Universal Robots PolyScope program: P1140 INVITE_training_1.urp

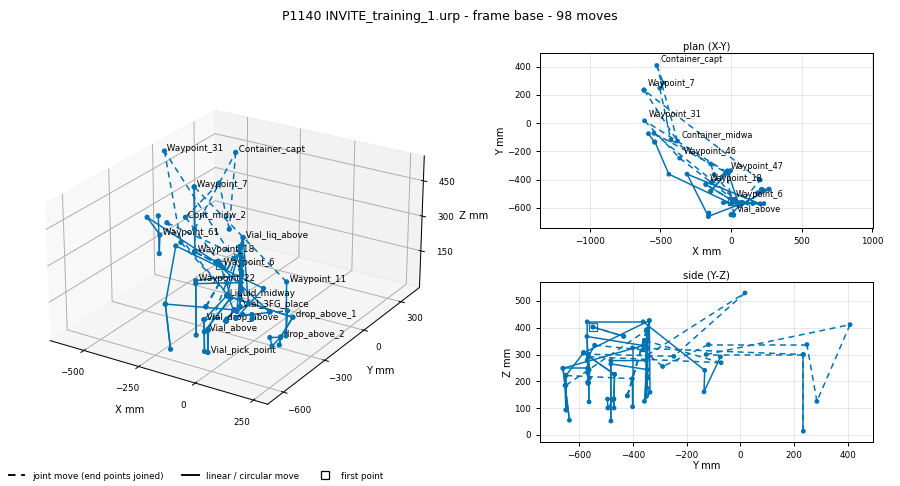
[picture p0: tool path of P1140 INVITE_training_1.urp in frame base, 98 of 125 moves have a stored position in this frame; points joined in program order, loops and branches not executed]
Program P1140 INVITE_training_1 (installation=default directory=/programs/02 Main Routines createdIn=5.10.1 lastSavedIn=5.19.0 robotSerialNumber=20245590068)
Calibrated DH parameters: a=[0.00013, -0.03651, -0.389144, 0.000102, 0.000008, 0]; d=[0.162613, 192.230671, -179.915756, -12.181517, 0.099698, 0.099535]; alpha=[1.57038, 0.002205, 0.004138, 1.570804, -1.571025, 0]; deltaTheta=[-0.000001, 1.484886, 4.928506, -0.130209, 0, 0]
InitVariablesNode variables(variable(name=AMR_Position, expression=struct(position_identifier=0, x1=0, x2=0, y1=0, y2=0, theta1=0, theta2=0)), variable(name=CAM_Pose, expression=p[0,0,0,0,0,0]), variable(name=CAM_Relation, expression=""), variable(name=CMD_Abort, expression=False), variable(name=CMD_Clear, expression=False), variable(name=CMD_Reset, expression=False), variable(name=CMD_Start, expression=False), variable(name=CMD_Suspend, expression=False), variable(name=CMD_Unhold, expression=False), variable(name=CMD_Unsuspend, expression=False), variable(name=CNT_Rack_Output, expression=0), variable(name=FNC_Freedrive, expression=False), variable(name=PRC_TubCounter, expression=0), variable(name=PRC_TubNumber, expression=0), variable(name=STP, expression=0), variable(name=TMR_Barcode, expression=0), variable(name=easyPickCount, expression=0), variable(name=easyPickCount_1, expression=0), variable(name=easyPickCount_2, expression=0), variable(name=easyPickCount_3, expression=0), variable(name=easyPickNoObj, expression=0), variable(name=easyPickNoObj_1, expression=0), variable(name=easyPickNoObj_2, expression=0), variable(name=easyPickNoObj_3, expression=0), variable(name=easyPickParts, expression=0), variable(name=easyPickParts_1, expression=0), variable(name=easyPickParts_2, expression=0), variable(name=easyPickParts_3, expression=0))
BeforeStart
  Folder Scripts
    Script file /programs/04 Scripts/001 SCRIPT Errors and Warnings Deifnes V0.2.script
      | #*****************************************************
      | # customer          :   UK Essen
      | # project name      :   P1132
      | #****************************************************
      | # controller        :
      | # software          :
      | #****************************************************
      | # author            :   E.Petrichenko
      | # Copyright (c)     :   United Robotics Group Health and Food GmbH
      | #                       An der Riede 2
      | #                       28816 Stuhr
      | #                       Germany
      | #****************************************************
      | # description       :   centrifuge actions for the application
      | # version:      	:   0.1
      | # created           :   22.08.2024
      | # updated           :
      | #****************************************************
      | # modifications     :
      | #
      | # date              :
      | # name              :
      | # reason            :
      | #****************************************************
      | 
      | 
      | #################################### VARIABLES DEFINITIONS ###################################
      | 
      | ERROR_POSE_NOT_REACHABLE = 1002
      | ERROR_ROBOT_ARM_NOT_IN_HOME_POSE = 1006
      | ERROR_NO_OBJECT_TO_PICK = 1010
      | ERROR_NOT_DOCKED = 2003
      | ERROR_NOT_REACHABLE_TARGET = 2007
      | ERROR_CHARGING_NOT_STARTED = 2008
      | ERROR_AMR_WRONG_MODE = 2009
      | ERROR_UNKNOWN_POSE = 2010
      | ERROR_NO_LANDMARK = 3002
      | ERROR_WRONG_ORDER = 4002
      | ERROR_CENTRIFUGE_CONNECTION = 5001
      | ERROR_CENTRIFUGE_POWER = 5002
      | ERROR_CENTRIFUGE = 5003
      | ERROR_CENTRIFUGE_LID = 5004
      | ERROR_CANNOT_OPEN_HATCH = 5006
      | ERROR_CANNOT_CLOSE_HATCH = 5008
      | ERROR_CANNOT_ROTATE = 5010
      | ERROR_CANNOT_START = 5011
      | ERROR_WRONG_KEY_POSE = 5012
      | ERROR_MISSIING_CENTRACK = 5013
      | 
      | WARNING_POSE_NOT_REACHABLE = 1002
      | WARNING_BATTERY_LEVEL = 2002
      | WARNING_NOT_REACHABLE_TARGET = 2007
      | 
      | 
      | ERROR = struct(
      |     FLAG = False,
      |     ID = 0,
      |     MSG = "")
      | 
      | WARNING = struct(
      |     FLAG = False,
      |     ID = 0,
      |     MSG = "")
      | 
      | 
      | #################################### FUNCTIONS ###################################
      | 
      | def set_error(error_id):
      |     ERROR.ID = error_id
      |     if (ERROR.ID == 0):
      |         ERROR.FLAG = False
      |         ERROR.MSG = ""
      |     else:
      |         ERROR.FLAG = True
      |         if(ERROR.ID == ERROR_POSE_NOT_REACHABLE):
      |             ERROR.MSG = "Pose is not reachable"
      |         elif(ERROR.ID == ERROR_NO_OBJECT_TO_PICK):
      |             ERROR.MSG = "No object to pick"
      |         elif(ERROR.ID == ERROR_NO_LANDMARK):
      |             ERROR.MSG = "No landmark detected"
      |         elif(ERROR.ID == ERROR_ROBOT_ARM_NOT_IN_HOME_POSE):
      |             ERROR.MSG = "Robot arm cannot go to home pose"
      |         elif(ERROR.ID == ERROR_AMR_WRONG_MODE):
      |             ERROR.MSG = "AMR is in the wrong mode"
      |         elif(ERROR.ID == ERROR_NOT_DOCKED):
      |             ERROR.MSG = "Could not dock to the charger"
      |         elif(ERROR.ID == ERROR_NOT_REACHABLE_TARGET):
      |             ERROR.MSG = "Could not reach the target"
      |         elif(ERROR.ID == ERROR_CHARGING_NOT_STARTED):
      |             ERROR.MSG = "Could not start charging"
      |         elif(ERROR.ID == ERROR_UNKNOWN_POSE):
      |             ERROR.MSG = "Unknown navigation target"
      |         elif(ERROR.ID == ERROR_CANNOT_OPEN_HATCH):
      |             ERROR.MSG = "Centrifuge Cannot open the hatch"
      |         elif(ERROR.ID == ERROR_CENTRIFUGE_CONNECTION):
      |             ERROR.MSG = "Cannot reach centrifuge"
      |         elif (ERROR.ID == ERROR_CANNOT_CLOSE_HATCH):
      |             ERROR.MSG = "Centrifuge Cannot close the hatch"
      |         elif (ERROR.ID == ERROR_CANNOT_START):
      |             ERROR.MSG = "Centrifuge Cannot start"
      |         elif (ERROR.ID == ERROR_CANNOT_ROTATE):
      |             ERROR.MSG = "Centrifuge Cannot rotate the rotor"
      |         elif (ERROR.ID == ERROR_WRONG_ORDER):
      |             ERROR.MSG = "Wrong parameter was recieved"
      |         elif (ERROR.ID == ERROR_CENTRIFUGE):
      |             ERROR.MSG = "Centrifuge is in Error"
      |         elif (ERROR.ID == ERROR_WRONG_KEY_POSE):
      |             ERROR.MSG = "Key is in the wrong position"
      |         elif(ERROR.ID == ERROR_MISSIING_CENTRACK):
      |             ERROR.MSG = "Missing rack for centrifuge set"
      |         elif(ERROR.ID == ERROR_CENTRIFUGE_POWER):
      |             ERROR.MSG = "Centrifuge is turned off"
      |         elif(ERROR.ID == ERROR_CENTRIFUGE_LID):
      |             ERROR.MSG = "Lid of the centrifuge is opened"
      |         else:
      |             ERROR.MSG = "Unknown code"
      |         end
      |         textmsg("ERROR:",ERROR)
      |     end
      | end
      | 
      | def set_warning(warning_id):
      |     WARNING.ID = warning_id
      |     if (WARNING.ID == 0):
      |         WARNING.FLAG = False
      |         WARNING.MSG = ""
      |     else:
      |         WARNING.FLAG = True
      |         if(WARNING.ID == WARNING_POSE_NOT_REACHABLE):
      |             WARNING.MSG = "Pose is not reachable"
      |         elif(WARNING.ID == WARNING_BATTERY_LEVEL):
      |             WARNING.MSG = "Batery level dropped to a certain level"
      |         elif(WARNING.ID == WARNING_NOT_REACHABLE_TARGET):
      |             WARNING.MSG = "Not reachable location of AMR"
      |         else:
      |             WARNING.MSG = "Unknown code"
      |         end
      |         textmsg("WARNING:",WARNING)
      |     end
      | end
      | 
      | 
      | def reset_error():
      |   ERROR.ID = 0
      |   ERROR.FLAG = False
      |   ERROR.MSG = ""
      | end
      | 
      | 
      | def reset_warning():
      |     WARNING.ID = 0
      |     WARNING.FLAG = False
      |     WARNING.MSG = ""
      |   end
    Script file /programs/04 Scripts/SCRIPT uGO V7.11.1.script
      | #*****************************************************
      | # customer          :
      | # project name      :   Standard Application
      | #****************************************************
      | # controller        :
      | # software          :
      | #****************************************************
      | # author            :   P. Koehnke
      | # Copyright (c)     :   United Robotics Group
      | #                       An der Riede 2
      | #                       28816 Stuhr
      | #                       Germany
      | #****************************************************
      | # description       :   interface for uGo
      | # version:      	:   6.0
      | # created           :   21.04.2022
      | # updated           :
      | #****************************************************
      | # modifications     :   add new rpc-functions to interchange more data
      | #
      | # date              :   2024-02-29
      | # name              :   P. Koehnke
      | # reason            :   implemtentation of PackML behavoiur in uGO
      | #****************************************************
      | #****************************************************
      | # modifications     :   add reflecting the UID of the uGO task back to uGO
      | #
      | # date              :   2024-07-02
      | # name              :   P. Koehnke
      | # reason            :   be sure to finish the right tasks
      | #****************************************************
      | 
      | # available rpc-functions:
      | #.on('con_check', (err, _params, callback) => callback(err, this.con_check()))
      | #.on('read_input', (err, params, callback) => callback(err, this.read_input(params[0], params[1])))
      | #.on('write_output', (err, params, callback) => callback(err, this.write_output(params[0], params[1], params[2])))
      | #.on('read_status', (err, params, callback) => callback(err, this.read_status(params[0])))
      | #.on('write_status', (err, params, callback) => callback(err, this.write_status(params[0], params[1])))
      | #.on('send_template', (err, params, callback) => callback(err, this.receive_state(params[0])))
      | #.on('receive_event', (err, params, callback) => callback(err, this.send_event()))
      | #.on('send_state', (err, params, callback) => callback(err, this.receive_state(params[0])))
      | #.on('send_error', (err, params, callback) => callback(err, this.receive_error(params[0])))
      | #.on('NotFound', (methodCalled, params) => LOG.warn('Method "', methodCalled, '" does not exist. ', { params }));
      | 
      | # =======================================================================
      | local IDX_CMD_STOP = 0
      | local IDX_CMD_RESET = 1
      | local IDX_CMD_START = 2
      | local IDX_CMD_HOLD = 3
      | local IDX_CMD_UNHOLD = 4
      | local IDX_CMD_SUSPEND = 5
      | local IDX_CMD_UNSUSPEND = 6
      | local IDX_CMD_ABORT = 7
      | local IDX_CMD_CLEAR = 8
      | local IDX_FNC_FREEDRIVE = 9
      | 
      | # uGo specific declarations
      | global UGO_Request_ID = ""
      | global UGO_UNIT_Task = ""
      | global UGO_Task_ID = 0
      | global UGO_Event = ""
      | local UGO_Enable_Control = False
      | local UGO = rpc_factory("xmlrpc", "http://192.168.12.120:8080")
      | local UGO_Ctrl_Cmd = [False, False, False, False, False, False, False, False, False, False]
      | 
      | local UGO_AMR_Pos = struct(position_identifier=0, x1=0, x2=0, y1=0, y2=0, theta1=0, theta2=0)
      | local UGO_EOAT = struct(object_picked=False)
      | 
      | def ugo_init(enable=True, rpc_address="http://192.168.12.120:8080"):
      |     # connection with uGo
      |     if enable:
      |         UGO = rpc_factory("xmlrpc", rpc_address)
      |         UGO_Enable_Control = True
      |     else:
      |         UGO_Enable_Control = False
      |     end
      | end
      | 
      | def ugo_event_controller():
      |     # interpret the given command and map it to the internal commands
      |     if UGO_Enable_Control:
      |         UGO_Event = UGO.receive_event()
      |     end
      | 
      |     UGO_Ctrl_Cmd[IDX_CMD_STOP] = (UGO_Event == "stop")
      |     UGO_Ctrl_Cmd[IDX_CMD_RESET] = (UGO_Event == "reset")
      |     UGO_Ctrl_Cmd[IDX_CMD_START] = (UGO_Event == "start")
      |     UGO_Ctrl_Cmd[IDX_CMD_HOLD] = (UGO_Event == "hold")
      |     UGO_Ctrl_Cmd[IDX_CMD_UNHOLD] = (UGO_Event == "un_hold")
      |     UGO_Ctrl_Cmd[IDX_CMD_SUSPEND] = (UGO_Event == "suspend")
      |     UGO_Ctrl_Cmd[IDX_CMD_UNSUSPEND] = (UGO_Event == "un_suspend")
      |     UGO_Ctrl_Cmd[IDX_CMD_ABORT] = (UGO_Event == "abort")
      |     UGO_Ctrl_Cmd[IDX_CMD_CLEAR] = (UGO_Event == "clear")
      |     UGO_Ctrl_Cmd[IDX_FNC_FREEDRIVE] = (UGO_Event == "freedrive")
      | 
      |     return UGO_Ctrl_Cmd
      | end
      | 
      | def ugo_translate_pml_state():
      |     # translate the current PML State to a string
      |     if (STATE == 1):
      |         return "STOPPING"
      |     elif (STATE == 2):
      |         return "STOPPED"
      |     elif (STATE == 3):
      |         return "RESETTING"
      |     elif (STATE == 4):
      |         return "IDLE"
      |     elif (STATE == 5):
      |         return "STARTING"
      |     elif (STATE == 6):
      |         return "EXECUTE"
      |     elif (STATE == 7):
      |         return "COMPLETING"
      |     elif (STATE == 8):
      |         return "COMPLETE"
      |     elif (STATE == 9):
      |         return "HOLDING"
      |     elif (STATE == 10):
      |         return "HELD"
      |     elif (STATE == 11):
      |         return "UNHOLDING"
      |     elif (STATE == 12):
      |         return "SUSPENDING"
      |     elif (STATE == 13):
      |         return "SUSPENDED"
      |     elif (STATE == 14):
      |         return "UNSUSPENDING"
      |     elif (STATE == 15):
      |         return "ABORTING"
      |     elif (STATE == 16):
      |         return "ABORTED"
      |     elif (STATE == 17):
      |         return "CLEARING"
      |     else:
      |         return "UNKNOWN"
      |     end
      | end
      | 
      | def ugo_update_outputs():
      |     #Update the outputs to uGo via xmplrpc service
      |     UGO.write_status("ROB_Skill", UGO_UNIT_Task)
      |     UGO.write_status("ROB_Battery", AMR_Battery)
      |     UGO.write_status("ROB_Gripper", OBJ_Picked)
      |     UGO.send_state(ugo_translate_pml_state(), UGO_UNIT_Task)
      |     UGO.send_error(ERROR.ID)
      |     #UGO.send_position(AMR_Position)
      | end
      | 
      | def ugo_get_task():
      |     # get the actual task to work on
      |     # added: reflecting the UID of the task back to uGO
      |     UGO_UNIT_Task = UGO.read_status("DSH_Workflow")
      |     if (UGO_UNIT_Task != ""):
      |         UGO_Request_ID = str_sub(UGO_UNIT_Task, 0, 39)
      |         UGO_Task_ID = to_num(str_sub(UGO_UNIT_Task, 40, 2))
      |         #ugo_tasks()
      |         return UGO_Task_ID
      |     else:
      |         return 0
      |     end
      | end
      | 
      | def ugo_pml_stopping():
      |     return True
      | end
      | 
      | def ugo_pml_resetting():
      |     ugo_get_task()
      |     if (UGO_UNIT_Task == ""):
      |         UGO_Request_ID = ""
      |         UGO_Task_ID = 0
      |         return True
      |     end
      |     return False
      | end
      | 
      | def ugo_pml_starting():
      |     #UGO_Task_Content = UGO.receive_task()
      |     return (UGO_UNIT_Task != "")
      | end
      | 
      | def ugo_pml_holding():
      |     return True
      | end
      | 
      | def ugo_pml_unholding():
      |     return True
      | end
      | 
      | def ugo_pml_suspending():
      |     return True
      | end
      | 
      | def ugo_pml_unsuspending():
      |     return True
      | end
      | 
      | def ugo_pml_completing():
      |     return True
      | end
      | 
      | def ugo_pml_aborting():
      |     return True
      | end
      | 
      | def ugo_pml_clearing():
      |     return True
      | end
      | 
      | # =======================================================================
      | # end of uGO script
      | # =======================================================================
    SuppressedNode
      Script file /programs/04 Scripts/SCRIPT Centrifuge Actions V0.3.script
        | #*****************************************************
        | # customer          :   UK Essen
        | # project name      :   P1132
        | #****************************************************
        | # controller        :
        | # software          :
        | #****************************************************
        | # author            :   E.Petrichenko
        | # Copyright (c)     :   United Robotics Group Health and Food GmbH
        | #                       An der Riede 2
        | #                       28816 Stuhr
        | #                       Germany
        | #****************************************************
        | # description       :   centrifuge actions for the application
        | # version:      	:   0.1
        | # created           :   22.08.2024
        | # updated           :
        | #****************************************************
        | # modifications     :
        | #
        | # date              :
        | # name              :
        | # reason            :
        | #****************************************************
        | 
        | 
        | #################################### VARIABLES DEFINITIONS ###################################
        | CNT_RESET_LOAD_TIMER = 60
        | CNT_Rotate_Error = False
        | CNT_Error = ""
        | CNT_LidState = 0
        | CNT_Timer_Start = 0
        | CNT_Timer_Counting = False
        | CNT_Hatch_State = 0
        | global CNT_State_Actual  = 0
        | CNT_KeyState = 0
        | Cent=rpc_factory("xmlrpc","http://192.168.12.125:50002")
        | 
        | ACTION_OPEN_HATCH = 5
        | ACTION_CLOSE_HATCH = 6
        | ACTION_START = 9
        | ACTION_INSPECT = 16
        | ACTION_ROTATE = 23
        | 
        | CNT_STATES_INIT = struct (
        |     UNSTARTABLE = 1,
        |     STOPPED = 2,
        |     STOPPED_UNSTARTABLE = 3,
        |     RUN_UP = 4,
        |     RUNNING = 8)
        | 
        | 
        | KEY_STATE_INIT = struct (
        |     TEACH = 1,
        |     LOCKED = 2,
        |     MIDDLE = 3)
        | 
        | LID_STATE_INIT = struct (
        |     CLOSED = 0,
        |     OPENED = 1)
        | #stopped_unstartable happens when lid or hatch is open
        | 
        | #################################### THREADS ###################################
        | 
        | thread Timer_CentThread():
        |     while (True):
        |         if (CNT_Timer_Counting):
        |             CNT_Timer_Start = CNT_Timer_Start + get_steptime()
        |         end
        |         sync()
        |     end
        | end
        | thread_timer_cent = run Timer_CentThread()
        | 
        | thread Cent_Thread():
        |     while (True):
        |         CNT_Hatch_State = Cent.hatchstate()
        |         CNT_State_Actual  = Cent.state()
        |         log_hatch_state(CNT_Hatch_State)
        |         log_centrifuge_state(CNT_State_Actual)
        |         sleep(0.5)
        |     end
        | end
        | run Cent_Thread()
        | 
        | #################################### FUNCTIONS ###################################
        | 
        | 
        | 
        | def cent_error_check():
        |     CNT_Error = Cent.geterror()
        |     CNT_KeyState = Cent.keystate()
        |     CNT_LidState = Cent.lidstate()
        | 
        |     if (CNT_Error == "88888888"):
        |         set_error(ERROR_CENTRIFUGE_POWER)
        |     elif (CNT_Error != "00000000"):
        |         set_error(ERROR_CENTRIFUGE)
        |         textmsg("CNT_Error:",CNT_Error)
        |     elif (CNT_KeyState != KEY_STATE_INIT.LOCKED):
        |         set_error(ERROR_WRONG_KEY_POSE)
        |     elif (CNT_LidState == LID_STATE_INIT.OPENED):
        |       set_error(ERROR_CENTRIFUGE_LID)
        |     end
        | 
        | end
        | 
        | 
        | def execute_cent_action(cent_action, cent_slot = 0):
        | 
        |     if (cent_action == ACTION_OPEN_HATCH):
        |         local cnt_hatch_moved = 0
        |         if (CNT_State_Actual  == 2):
        |             cnt_hatch_moved = Cent.move_hatch(2)
        |             if (cnt_hatch_moved == -1):
        |                 set_error(ERROR_CANNOT_OPEN_HATCH)
        |             end
        |         elif (CNT_State_Actual  == 3):
        |             textmsg("WARNING: Centrifuge is already opened", True)
        |         else:
        |             set_error(ERROR_WRONG_ORDER)
        |             textmsg("ERROR: Centrifuge state is not corresponded with the required task", True)
        |         end
        | 
        |     elif (cent_action == ACTION_CLOSE_HATCH):
        |         cnt_hatch_moved = Cent.move_hatch(1)
        |         if (cnt_hatch_moved == -1):
        |             set_error(ERROR_CANNOT_CLOSE_HATCH)
        |         end
        | 
        |     elif (cent_action == ACTION_START):
        |         Cent.start()
        |         CNT_Timer_Start = 0
        |         CNT_Timer_Counting = True
        |         while ((CNT_State_Actual  != CNT_STATES_INIT.RUN_UP and CNT_State_Actual  != CNT_STATES_INIT.RUNNING) and CNT_Timer_Start < CNT_RESET_LOAD_TIMER and not CMD_Stop and not CMD_Hold):
        |             sleep(0.5)
        | 
        |         end
        | CNT_Timer_Counting = False
        |         if (CNT_Timer_Start >= CNT_RESET_LOAD_TIMER ):
        |             set_error(ERROR_CANNOT_START)
        |             if (CNT_State_Actual == CNT_STATES_INIT.UNSTARTABLE or CNT_State_Actual == CNT_STATES_INIT.STOPPED_UNSTARTABLE):
        |                 set_error(ERROR_WRONG_ORDER)
        |                 textmsg("ERROR: Centrifuge state is not corresponded with the required task", True)
        |             end
        |         end
        |     elif (cent_action == ACTION_INSPECT):
        |         if (CNT_Rotate_Error == False):
        |             set_error(ERROR_CANNOT_ROTATE)
        |         else:
        |             CNT_Rotate_Error = Cent.posreached(6 *(cent_slot-1) + 1)
        |             if (CNT_Rotate_Error == False):
        |               set_error(ERROR_CANNOT_ROTATE)
        |             end
        |         end
        | 
        | 
        |     elif (cent_action == ACTION_ROTATE):
        |         CNT_Rotate_Error = False
        |         CNT_Rotate_Error = Cent.move_rotor(6 *(cent_slot-1) + 1)
        |         return CNT_Rotate_Error
        |     else:
        |         set_error(ERROR_WRONG_ORDER)
        |     end
        | end
    Script file /programs/04 Scripts/SCRIPT PackML V1.2.1.script
      | # PackML
      | 
      | IO_ADDRESS_CMD_STOP = 1
      | IO_ADDRESS_CMD_RESET = 7
      | IO_ADDRESS_CMD_START = 0
      | 
      | EXT_ADDRESS_CMD_STOP = 0
      | EXT_ADDRESS_CMD_RESET = 1
      | EXT_ADDRESS_CMD_START = 2
      | EXT_ADDRESS_CMD_HOLD = 3
      | EXT_ADDRESS_CMD_UNHOLD = 4
      | EXT_ADDRESS_CMD_SUSPEND = 5
      | EXT_ADDRESS_CMD_UNSUSPEND = 6
      | EXT_ADDRESS_CMD_ABORT = 7
      | EXT_ADDRESS_CMD_CLEAR = 8
      | EXT_ADDRESS_FNC_FREEDRIVE = 9
      | 
      | global EXT_CtrlCmd = [False, False, False, False, False, False, False, False, False, False]
      | 
      | EXT_Control_by = "uGO"
      | 
      | global CMD_Abort = False
      | global CMD_Clear = False
      | global CMD_Stop = False
      | global CMD_Reset = False
      | global CMD_Start = False
      | global CMD_Hold = False
      | global CMD_Unhold = False
      | global CMD_Suspend = False
      | global CMD_Unsuspend = False
      | global FNC_Freedrive = False
      | 
      | CND_Suspend = False         # condition for suspend command
      | CND_Unsuspend = False       # condition for unsuspend command
      | 
      | thread Get_Pml_Command():
      |     while (True):
      |         if (EXT_Control_by == "uGO"):
      |             EXT_CtrlCmd = ugo_event_controller()
      |         elif (EXT_Control_by == "Leitsystem"):
      |             # EXT_CtrlCmd = Leitsystem
      |         end
      |         # ---------- Abort ---------- #
      |         if ((not STATE == 15) and (not STATE == 16) and EXT_CtrlCmd[EXT_ADDRESS_CMD_ABORT]):
      |             CMD_Abort = True
      |             CMD_Stop = False
      |         elif ((STATE == 17) and not EXT_CtrlCmd[EXT_ADDRESS_CMD_ABORT]):
      |             CMD_Abort = False
      |         end
      |         # ---------- Stop ---------- #
      |         if ((not STATE == 1) and (not STATE == 2) and (get_standard_digital_in(IO_ADDRESS_CMD_STOP) or EXT_CtrlCmd[EXT_ADDRESS_CMD_STOP])):
      |             CMD_Stop = True
      |             if get_standard_digital_in(IO_ADDRESS_CMD_STOP):
      |                 log_state("Stop command by pushbutton")
      |             elif EXT_CtrlCmd[EXT_ADDRESS_CMD_STOP]:
      |                 log_state("Stop command by external control")
      |             end
      |         elif (STATE == 2) and (not get_standard_digital_in(IO_ADDRESS_CMD_STOP)) and (not EXT_CtrlCmd[EXT_ADDRESS_CMD_STOP]):
      |             CMD_Stop = False
      |         end
      |         CMD_Hold = (STATE == 6 or STATE == 10) and not CMD_Stop and (ERROR.FLAG or EXT_CtrlCmd[EXT_ADDRESS_CMD_HOLD])
      |         CMD_Reset = (STATE == 2 or STATE == 8) and not CMD_Stop and (read_input_boolean_register(5) or EXT_CtrlCmd[EXT_ADDRESS_CMD_RESET])
      |         CMD_Start = (STATE == 4) and not CMD_Stop and (get_standard_digital_in(IO_ADDRESS_CMD_START) or EXT_CtrlCmd[EXT_ADDRESS_CMD_START])
      |         CMD_Unhold = (STATE == 10) and not CMD_Stop and (get_standard_digital_in(IO_ADDRESS_CMD_START) or EXT_CtrlCmd[EXT_ADDRESS_CMD_UNHOLD])
      |         CMD_Suspend = (STATE == 6) and not CMD_Stop and (CND_Suspend or EXT_CtrlCmd[EXT_ADDRESS_CMD_SUSPEND])
      |         CMD_Unsuspend = (STATE == 13) and not CMD_Stop and (CND_Unsuspend or EXT_CtrlCmd[EXT_ADDRESS_CMD_UNSUSPEND])
      |         CMD_Clear = (STATE == 16) and EXT_CtrlCmd[EXT_ADDRESS_CMD_CLEAR]
      |         FNC_Freedrive = (STATE == 10) and EXT_CtrlCmd[EXT_ADDRESS_FNC_FREEDRIVE]
      |         sleep(0.1)
      |     end
      | end
      | 
      | thread_pml_command_handler = run Get_Pml_Command()
      | 
      | def command_manager(external_control="uGO", cond_suspend=False, cond_unsuspend=False):
      | 
      |     EXT_Control_by = external_control
      |     CND_Suspend = cond_suspend
      |     CND_Unsuspend = cond_unsuspend
      | 
      |     if (CMD_Abort and STATE != 15 and STATE != 16):
      |         STATE = 15
      |     elif (CMD_Stop and STATE != 1 and STATE != 2):
      |         STATE = 1
      |     end
      |     return False
      | end
      | 
      | def stopping():
      |     if (EXT_Control_by == "uGO"):
      |         return ugo_pml_stopping()
      |     elif (EXT_Control_by == "Leitsystem"):
      |         # EXT_CtrlCmd = Leitsystem
      |     else:
      |         return True
      |     end
      |     return False
      | end
      | 
      | def resetting():
      |     if (EXT_Control_by == "uGO"):
      |         return ugo_pml_resetting()
      |     elif (EXT_Control_by == "Leitsystem"):
      |         # EXT_CtrlCmd = Leitsystem
      |     else:
      |         return True
      |     end
      |     return False
      | end
      | 
      | def starting():
      |     if (EXT_Control_by == "uGO"):
      |         return ugo_pml_starting()
      |     elif (EXT_Control_by == "Leitsystem"):
      |         # EXT_CtrlCmd = Leitsystem
      |     else:
      |         return True
      |     end
      |     return False
      | end
      | 
      | def holding():
      |     if (EXT_Control_by == "uGO"):
      |         return ugo_pml_holding()
      |     elif (EXT_Control_by == "Leitsystem"):
      |         # EXT_CtrlCmd = Leitsystem
      |     else:
      |         return True
      |     end
      |     return False
      | end
      | 
      | def unholding():
      |     if (EXT_Control_by == "uGO"):
      |         return ugo_pml_unholding()
      |     elif (EXT_Control_by == "Leitsystem"):
      |         # EXT_CtrlCmd = Leitsystem
      |     else:
      |         return True
      |     end
      |     return False
      | end
      | 
      | def suspending():
      |     if (EXT_Control_by == "uGO"):
      |         return ugo_pml_suspending()
      |     elif (EXT_Control_by == "Leitsystem"):
      |         # EXT_CtrlCmd = Leitsystem
      |     else:
      |         return True
      |     end
      |     return False
      | end
      | 
      | def unsuspending():
      |     if (EXT_Control_by == "uGO"):
      |         return ugo_pml_unsuspending()
      |     elif (EXT_Control_by == "Leitsystem"):
      |         # EXT_CtrlCmd = Leitsystem
      |     else:
      |         return True
      |     end
      |     return False
      | end
      | 
      | def completing():
      |     if (EXT_Control_by == "uGO"):
      |         return ugo_pml_completing()
      |     elif (EXT_Control_by == "Leitsystem"):
      |         # EXT_CtrlCmd = Leitsystem
      |     else:
      |         return True
      |     end
      |     return False
      | end
      | 
      | def aborting():
      |     if (EXT_Control_by == "uGO"):
      |         return ugo_pml_aborting()
      |     elif (EXT_Control_by == "Leitsystem"):
      |         # EXT_CtrlCmd = Leitsystem
      |     else:
      |         return True
      |     end
      |     return False
      | end
      | 
      | def clearing():
      |     if (EXT_Control_by == "uGO"):
      |         return ugo_pml_clearing()
      |     elif (EXT_Control_by == "Leitsystem"):
      |         # EXT_CtrlCmd = Leitsystem
      |     else:
      |         return True
      |     end
      |     return False
      | end
    Script file /programs/04 Scripts/SCRIPT Utility V5.5.script
      | #*****************************************************
      | # customer          :   tbd
      | # project name      :   tbd
      | #****************************************************
      | # controller        :
      | # software          :
      | #****************************************************
      | # author            :   P. Koehnke (+49 1628859904; p.koehnke@unitedrobotics.group)
      | # Copyright (c)     :   United Robotics Group Health and Food GmbH
      | #                       An der Riede 2
      | #                       28816 Stuhr
      | #                       Germany
      | #****************************************************
      | # description       :   utility programs for the application
      | # version:      	:   3.1
      | # created           :   30.01.2023
      | # updated           :
      | #****************************************************
      | # modifications     :   get_tool_free_pose_2(), get_index_from_list()
      | #
      | # date              :   05.01.2024
      | # name              :   PK
      | # reason            :
      | #****************************************************
      | 
      | def found_in_matrix(data, req_id, req_idx):
      |     local id = -1
      |     local dimensions = size(data)
      |     local loop_dataset = 0
      | 
      |     while (id != req_id and loop_dataset < dimensions[0]):
      |         id = data[loop_dataset, 0]
      |         if (id == req_id):
      |             return data[loop_dataset, req_idx]
      |         else:
      |             loop_dataset = loop_dataset + 1
      |         end
      |     end
      | end
      | 
      | def found_in_list(value, list):
      |     local idx = 0
      | 
      |     while (idx < length(list)):
      |         if (value == list[idx]):
      |             return True
      |         end
      |         idx = idx + 1
      |     end
      |     return False
      | end
      | 
      | def get_index_from_list(list, value = -1):
      |     local idx = 0
      | 
      |     while (idx < length(list)):
      |         if (value == -1):
      |             if (list[idx] != 0):
      |                 return idx
      |             end
      |         else:
      |             if (list[idx] == value):
      |                 return idx
      |             end
      |         end
      |         idx = idx + 1
      |     end
      |     return -1
      | end
      | 
      | def find_object_by_type(list, type=0):
      |     local object = list[0]
      |     local i = 0
      | 
      |     while i < length(list):
      |         object = list[i]
      |         if object.type == type:
      |             return object
      |         end
      |         i = i + 1
      |     end
      | end
      | 
      | def pose_RPY2RotVec(pose):
      |     local rotvec = rpy2rotvec([d2r(pose[3]), d2r(pose[4]), d2r(pose[5])])
      |     return p[pose[0], pose[1], pose[2], rotvec[0], rotvec[1], rotvec[2]]
      | end
      | 
      | def pose_RotVec2RPY(pose):
      |     local rpy = rotvec2rpy([pose[3], pose[4], pose[5]])
      |     return p[pose[0], pose[1], pose[2], r2d(rpy[0]), r2d(rpy[1]), r2d(rpy[2])]
      | end
      | 
      | def swivel(frame_ref, angles = [0, 0, 0], pose = p[0, 0, 0, 0, 0, 0]):
      | 
      |     local rpy_ref = [0, 0, 0]
      |     local rpy_new = [0, 0, 0]
      |     local rotvec_new = [0, 0, 0]
      |     local pose_from = p[0, 0, 0, 0, 0, 0]
      |     local pose_to = p[0, 0, 0, 0, 0, 0]
      |     local i = 0
      | 
      |     if (pose == p[0, 0, 0, 0, 0, 0]):
      |         pose_to = pose_trans(pose_inv(frame_ref), get_actual_tcp_pose())
      |     else:
      |         pose_to = pose
      |     end
      | 
      |     rpy_ref = rotvec2rpy(frame_ref[3], frame_ref[4], frame_ref[5])
      | 
      |     while (i < 3):
      |         rpy_new[i] = rpy_ref[i] + d2r(angles[i])
      |         i = i + 1
      |     end
      | 
      |     rotvec_new = rpy2rotvec(rpy_new)
      |     pose_from = p[0, 0, 0, rotvec_new[0], rotvec_new[1], rotvec_new[2]]
      |     pose_to = p[pose_to[0], pose_to[1], pose_to[2], rotvec_new[0], rotvec_new[1], rotvec_new[2]]
      | 
      |     return pose_trans(pose_from, pose_to)
      | end
      | 
      | def get_random_pose(pose_ref, mode = "", range_max = [0, 0, 0]):
      |     # modi: "cubic", "rotation"
      |     # getting a random pose in the x/y-plane. range can be set for each
      |     # translation and rotation.
      |     local rpy_random = [0, 0, 0]
      |     local rotvec_random = [0, 0, 0]
      |     local pose_random = pose_ref
      |     local i = 0
      | 
      |     if (mode == "cubic"):
      |         # cubic mode: random pose takes only x, y and z
      |         i = 0
      |         while (i < 3):
      |             pose_random[i] = pose_ref[i] + range_max[i] * (random() - 0.5)
      |             i = i + 1
      |         end
      |         return pose_random
      | 
      |     elif (mode == "rotation"):
      |         i = 0
      |         while (i < 3):
      |             rpy_random[i] = d2r(range_max[i]) * (random() - 0.5)
      |             i = i + 1
      |         end
      |         rotvec_random = rpy2rotvec(rpy_random)
      |         pose_random = pose_trans(p[0, 0, 0, rotvec_random[0], rotvec_random[1], rotvec_random[2]], pose_ref)
      |         return pose_random
      | 
      |     else:
      |         # unknown mode, return pose_ref
      |         return pose_ref
      |     end
      | end
      | 
      | def get_pattern_pos_rectangle(counter, direction, pattern, patterninc = [0, 0], patternsize = [0, 0]):
      |     # defines the position inside a rectangular pattern
      |     # pattern describes, how many objects are in x-direction and how many in y-direction [x, y]
      |     # patternsize will give the total length of each direction [x, y]
      |     local X_Fac = 0
      |     local Y_Fac = 0
      |     local max = pattern[0] * pattern[1]
      |     local i = 0
      | 
      |     if (1 > counter or counter > max):
      |         counter = 1
      |     end
      | 
      |     if pattern[0] == 0:
      |         pattern[0] = 1
      |     end
      | 
      |     if pattern[1] == 0:
      |         pattern[1] = 1
      |     end
      | 
      |     if (direction == "Y" or direction == "y"):
      |         X_Fac = floor((counter - 1) / pattern[1])
      |         Y_Fac = (counter - 1) % pattern[1]
      |     elif (direction == "X" or direction == "x"):
      |         X_Fac = (counter - 1) % pattern[0]
      |         Y_Fac = floor((counter - 1) / pattern[0])
      |     end
      | 
      |     if patternsize != [0, 0]:
      |         while i < 2:
      |             if pattern[i] > 1:
      |                 patterninc[i] = patternsize[i] / (pattern[i] - 1)
      |             end
      |             i = i + 1
      |         end
      |     end
      | 
      |     return p[X_Fac * patterninc[0], Y_Fac * patterninc[1], 0, 0, 0, 0]
      | end
      | 
      | def get_pattern_pos_circle(counter, radius, angle, direction, pattern, patternsize = [0, 0]):
      |     # get the patternpos for a circular pattern through a counter
      |     # need the radius and the angle in radiants
      |     local X_Fac = 0
      |     local Y_Fac = 0
      |     local rad_bow = 0
      |     local radius_cal = 0
      |     local ref = p[0, 0, 0, 0, 0, 0]
      | 
      |     if pattern[0] == 0:
      |         pattern[0] = 1
      |     end
      | 
      |     if pattern[1] == 0:
      |         pattern[1] = 1
      |     end
      | 
      |     if (direction == "Y" or direction == "y"):
      |         X_Fac = floor((counter - 1) / pattern[1])
      |         Y_Fac = (counter - 1) % pattern[1]
      |     elif (direction == "X" or direction == "x"):
      |         X_Fac = (counter - 1) % pattern[0]
      |         Y_Fac = floor((counter - 1) / pattern[0])
      |     end
      | 
      |     # the opening angle will be calculated in x-direction
      |     # works only between -90 and 90 degree
      |     if pattern[0] > 1:
      |         rad_bow = - angle / (pattern[0] - 1) * X_Fac + angle / 2
      |     end
      | 
      |     if (counter % 2 == 0 and pattern[1] > 1):
      |         radius_cal = radius - patternsize[1] / (pattern[1])
      |     else:
      |         radius_cal = radius + patternsize[1] / (pattern[1])
      |     end
      |     ref = p[0, radius_cal, 0, 0, 0, 0]
      | 
      |     return p[ref[0] * cos(rad_bow) - ref[1] * sin(rad_bow), (ref[0] * sin(rad_bow) + ref[1] * cos(rad_bow)) - radius, 0, 0, 0, 0]
      | end
      | 
      | def get_pattern_counter(pose, direction, pattern, patterninc = [0, 0], patternsize = [0, 0]):
      |     # returns the counter for a pattern from a given cartesian pose
      |     local patternpose = p[pose[0], pose[1], 0, 0, 0, 0]
      |     local X_Fac = 0
      |     local Y_Fac = 0
      |     local i = 0
      | 
      |     if patternsize != [0, 0]:
      |         while i < 2:
      |             if pattern[i] > 1:
      |                 patterninc[i] = patternsize[i] / (pattern[i] - 1)
      |             else:
      |                 pattern[i] = 0
      |             end
      |             i = i + 1
      |         end
      |     end
      | 
      |     # calculation of the counter in the desired axis-direction
      |     if (direction == "x" or direction == "X"):
      |         if patterninc[0] > 0:
      |             X_Fac = ceil((patternpose[0] + patterninc[0] / 2) / patterninc[0])
      |             if X_Fac < 0:
      |                 X_Fac = 0
      |             end
      |         end
      |         if patterninc[1] > 0:
      |             Y_Fac = floor((patternpose[1] + patterninc[1] / 2) / patterninc[1])
      |             if Y_Fac < 0:
      |                 Y_Fac = 0
      |           end
      |         end
      |         return Y_Fac * pattern[0] + X_Fac
      |     elif (direction == "y" or direction == "Y"):
      |         if patterninc[0] > 0:
      |             X_Fac = floor((patternpose[0] + patterninc[0] / 2) / patterninc[0])
      |         end
      |         if patterninc[1] > 0:
      |             Y_Fac = ceil((patternpose[1] + patterninc[1] / 2) / patterninc[1])
      |         end
      |         return X_Fac * pattern[1] + Y_Fac
      |     end
      | end
      | 
      | def get_plc_reg(mod_sig_name):
      |     return integer_to_binary_list(modbus_get_signal_status(mod_sig_name))
      | end
      | 
      | def set_plc_reg(mod_sig_name, mod_sig_list):
      |     modbus_set_output_register(mod_sig_name, binary_list_to_integer(mod_sig_list), False)
      | end
      | 
      | def check_decapping(offset = 0, timeout = 5, abort = False):
      |     # checken, ob der Deckel schon ab ist
      |     local start = get_actual_tcp_pose()
      |     local current_offset = 0
      |     local timecounter = 0
      |     while (current_offset < offset and not abort):
      |         current_offset = pose_dist(start, get_actual_tcp_pose())
      |         timecounter = timecounter + 1
      |         if (timecounter * 0.5 == timeout):
      |             break
      |         end
      |         sleep(0.5)
      |     end
      |     stopl(0.5)
      | end
      | 
      | def check_capping(torque = 0):
      |     # checken, wann der Deckel verschraubt ist
      |     force_mode(get_actual_tcp_pose(), [0, 0, 1, 0, 0, 0], [0, 0, -2.0, 0, 0, 0], 2, [0.01, 0.01, 0.001, 0.01, 0.01, 0.01])
      | end
      | 
      | def is_reachable(frame, poses, offsets = [0, 0, 0]):
      |     local idx = 0
      |     local pose = p[0, 0, 0, 0, 0, 0]
      | 
      |     while (idx < length(poses)):
      |         pose = poses[idx]
      |         pose[0] = pose[0] + offsets[0]
      |         pose[1] = pose[1] + offsets[1]
      |         pose[2] = pose[2] + offsets[2]
      | 
      |         if pose != p[0, 0, 0, 0, 0, 0]:
      |             if (not get_inverse_kin_has_solution(pose_trans(frame, pose))):
      |                 textmsg(str_cat(str_cat("Pose ", to_str(idx + 1)), " is not reachable"))
      |                 return False
      |             end
      |         end
      |         idx = idx + 1
      |     end
      |     return True
      | end
      | 
      | def is_within_limits(frame, poses, offsets = [0, 0, 0]):
      |     local idx = 0
      |     local pose = p[0, 0, 0, 0, 0, 0]
      | 
      |     while (idx < length(poses)):
      |         pose = poses[idx]
      |         pose[0] = pose[0] + offsets[0]
      |         pose[1] = pose[1] + offsets[1]
      |         pose[2] = pose[2] + offsets[2]
      | 
      |         if is_reachable(frame = frame, poses = poses, offsets = offsets):
      |             if (not is_within_safety_limits(get_inverse_kin(pose_trans(frame, pose), get_actual_joint_positions()))):
      |                 textmsg(str_cat(str_cat("Pose ", to_str(idx + 1)), "is out of joint limits"))
      |                 return False
      |             else:
      |                 idx = idx + 1
      |             end
      |         else:
      |             return False
      |         end
      |     end
      |     return True
      | end
      | 
      | 
      | def string_to_list(string, separator = "," , endDelimiter = ";" , capacity = 50):
      |     local string_length = str_len(string)
      |     local list_out = make_list(length = elements_in_string(string), initial_value = -1, capacity = capacity)
      |     local cnt = 0
      |     local idx = 0
      | 
      |     while cnt < string_length-1 :
      |       textmsg("new loop")
      |       textmsg(to_str(idx))
      |       local sepAt = str_find(string, separator, cnt)
      |       textmsg(to_str(sepAt))
      |       if sepAt < 0 :
      |           sepAt = str_find(string, endDelimiter, cnt)
      |       end
      |       list_out[idx] = to_num(str_sub(string, cnt, sepAt-cnt))
      |       idx = idx +1
      |       cnt = sepAt + 1
      |     end
      | 
      |     return list_out
      | end
      | 
      | def elements_in_string(string, separator = "," , endDelimiter = ";" , capacity = 50):
      |    local string_length = str_len(string)
      |     local len = 0
      |     local sepAt = 0
      | 
      |     while sepAt < string_length-1 and sepAt>=0 :
      |       local sepAt = str_find(string, separator, sepAt+1)
      |       len = len +1
      |     end
      | 
      |     return len
      | end
    Script file /programs/04 Scripts/SCRIPT uML Lights V1.2.script
      | #****************************************************
      | # product           : uLabMobile
      | # language          : urscript
      | #****************************************************
      | # author            :   D.Kreugel
      | # Copyright (c)     :   United Robotics Group
      | #                       An der Riede 2
      | #                       28816 Stuhr
      | #                       Germany
      | #****************************************************
      | # description       :   led controls for uLabMobile
      | # version:      	:   1.2
      | # created           :   09.08.2024
      | # updated           :
      | #****************************************************
      | # modifications     :   changed conditions to switch lights (not only pml state but also charging state)
      | #
      | # date              :   09.08.2024
      | # name              :   PK
      | # reason            :   due to the change in project P1117, we run to often through every state. This leads to to much colorchanges
      | #****************************************************
      | 
      | # HARDWARE CONFIGURATION
      | LED_GREEN = struct(type="CO",id=5)
      | LED_RED = struct(type="CO",id=6)
      | LED_BLUE = struct(type="CO",id=7)
      | 
      | def set_output(type,id,state=True):
      |     if(type=="CO"):
      |         set_configurable_digital_out(id,state)
      |     elif(type=="DO"):
      |         set_standard_digital_out(id,state)
      |     end
      | end
      | 
      | def led_red_on():
      |     set_output(LED_RED.type,LED_RED.id,True)
      | end
      | 
      | def led_red_off():
      |     set_output(LED_RED.type,LED_RED.id,False)
      | end
      | 
      | def led_green_on():
      |     set_output(LED_GREEN.type,LED_GREEN.id,True)
      | end
      | 
      | def led_green_off():
      |     set_output(LED_GREEN.type,LED_GREEN.id,False)
      | end
      | 
      | def led_blue_on():
      |     set_output(LED_BLUE.type,LED_BLUE.id,True)
      | end
      | 
      | def led_blue_off():
      |     set_output(LED_BLUE.type,LED_BLUE.id,False)
      | end
      | 
      | 
      | # COLOR MIX
      | def color_blue():
      |     led_blue_on()
      |     led_green_off()
      |     led_red_off()
      | end
      | 
      | def color_red():
      |     led_blue_off()
      |     led_green_off()
      |     led_red_on()
      | end
      | 
      | def color_green():
      |     led_blue_off()
      |     led_green_on()
      |     led_red_off()
      | end
      | 
      | def color_yellow():
      |     led_blue_off()
      |     led_green_on()
      |     led_red_on()
      | end
      | 
      | def color_lightblue():
      |     led_blue_on()
      |     led_green_on()
      |     led_red_off()
      | end
      | 
      | def color_violet():
      |     led_blue_on()
      |     led_green_off()
      |     led_red_on()
      | end
      | 
      | def color_white():
      |     led_blue_on()
      |     led_green_on()
      |     led_red_on()
      | end
      | 
      | def led_off():
      |     led_blue_off()
      |     led_green_off()
      |     led_red_off()
      | end
      | 
      | # COLOR FOR STATES
      | thread Thread_Lights():
      |     while(True):
      |         # Stopping
      |         if (STATE == 1):
      |             color_red()
      |             sleep(0.5)
      |             led_off()
      |         # Stopped
      |         elif (STATE == 2):
      |             color_red()
      |         # Resetting
      |         # elif (STATE == 3):
      |         #     color_white()
      |         #     sleep(0.5)
      |         #     led_off()
      |         # Idle
      |         elif (AMR_Charging):
      |             color_white()
      |         # Starting
      |         # elif (STATE == 5):
      |         #     color_lightblue()
      |         #     sleep(0.5)
      |         #     led_off()
      |         # Execute
      |         # elif (STATE == 6):
      |         #     color_lightblue()
      |         # Completing
      |         # elif (STATE == 7):
      |         #     color_green()
      |         #     sleep(0.5)
      |         #     led_off()
      |         # # Complete
      |         # elif (STATE == 8):
      |         #     color_green()
      |         # Holding
      |         elif (STATE == 9):
      |             color_red()
      |             sleep(0.5)
      |             led_off()
      |         # Held
      |         elif (STATE == 10):
      |             color_red()
      |         # Unholding
      |         elif (STATE == 11):
      |             color_yellow()
      |             sleep(0.5)
      |             led_off()
      |         # Suspending
      |         elif (STATE == 12):
      |             color_blue()
      |             sleep(0.5)
      |             led_off()
      |         # Suspended
      |         elif (STATE == 13):
      |             color_blue()
      |         # Unsuspending
      |         elif (STATE == 14):
      |             color_yellow()
      |             sleep(0.5)
      |             led_off()
      |         # Aborting
      |         elif (STATE == 15):
      |             color_red()
      |             sleep(0.5)
      |             led_off()
      |         # Aborted
      |         elif (STATE == 16):
      |             color_red()
      |         # Clearing
      |         elif (STATE == 17):
      |             color_yellow()
      |             sleep(0.5)
      |             led_off()
      |         else:
      |             color_lightblue()
      |         end
      |         sleep(0.5)
      |     end
      | end
      | 
      | thread_lights_handler = run Thread_Lights()
    Script file /programs/04 Scripts/SCRIPT Transitions V8.0.script
      | #*****************************************************
      | # customer          :   INTERNAL
      | # project name      :
      | #****************************************************
      | # controller        :   UR
      | # software          :   5.13
      | #****************************************************
      | # author            :   P. Koehnke
      | # Copyright (c)     :   United Robotics Group
      | #                       An der Riede 2
      | #                       28816 Stuhr
      | #                       Germany
      | #****************************************************
      | # description       :   transition between workareas
      | # version:      	:   1.2
      | # created           :   28.02.2024
      | # updated           :
      | #****************************************************
      | # modifications     :
      | #
      | # date              :
      | # name              :
      | # reason            :
      | #****************************************************
      | 
      | ######################### further development #########################
      | #   - that the robot can switch the configuration, if necessary
      | #   - introduction of structs
      | #######################################################################
      | 
      | ######################### to be adjusted #########################
      | 
      | local WORKAREA_1 = [-0.280,-0.680,-0.001, 0.280, 0.100, 1.000]    # workarea 1 (platform)
      | local WORKAREA_2 = [-1.000,-1.000,-1.000,-0.280, 0.100, 1.000]    # workarea 2 (front right)
      | local WORKAREA_3 = [-1.000, 0.100,-1.000, 0.000, 1.000, 1.000]    # workarea 3 (back right)
      | local WORKAREA_4 = [ 0.000, 0.100,-1.000, 1.000, 1.000, 1.000]    # workarea 4 (back left)
      | local WORKAREA_5 = [ 0.280,-1.000,-1.000, 1.000, 0.100, 1.000]    # workarea 5 (front left)
      | local WORKAREA_6 = [-0.280,-1.000,-1.000, 0.280,-0.680, 1.000]    # workarea 6 (front front)
      | local WORKAREA_7 = [0,0,0,0,0,0]    # reserved
      | local WORKAREA_8 = [0,0,0,0,0,0]    # reserved
      | local WORKAREA_9 = [0,0,0,0,0,0]    # reserved
      | local WORKAREA_10 = [0,0,0,0,0,0]   # reserved
      | 
      | local PSE_WA_1 = p[ 0.000,-0.450, 0.300, 0.000, 0.000, 0.000]
      | local PSE_WA_2 = p[-0.300,-0.300, 0.300, 0.000, 0.000, d2r(-90)]
      | local PSE_WA_3 = p[-0.300, 0.300, 0.300, 0.000, 0.000, d2r(-135)]
      | local PSE_WA_4 = p[ 0.300, 0.300, 0.300, 0.000, 0.000, d2r(135)]
      | local PSE_WA_5 = p[ 0.300,-0.300, 0.300, 0.000, 0.000, d2r(90)]
      | local PSE_WA_6 = p[ 0.000,-0.600, 0.300, 0.000, 0.000, 0.000]       # reserved
      | local PSE_WA_7 = p[ 0.000, 0.000, 0.000, 0.000, 0.000, 0.000]       # reserved
      | local PSE_WA_8 = p[ 0.000, 0.000, 0.000, 0.000, 0.000, 0.000]       # reserved
      | local PSE_WA_9 = p[ 0.000, 0.000, 0.000, 0.000, 0.000, 0.000]       # reserved
      | local PSE_WA_10 = p[ 0.000, 0.000, 0.000, 0.000, 0.000, 0.000]      # reserved
      | 
      | global JNT_HOME = [-1.23163,-1.29627,-1.86552,-1.55102, 1.57761, 1.910]
      | local JNT_STANDARD_C1 = [ 1.57,-1.57, 1.57,-1.57,-1.57,0]
      | local JNT_STANDARD_C2 = [-1.57,-1.57,-1.57,-1.57, 1.57,0]
      | local ANGLE_MIN_DEG = -110
      | local ANGLE_MAX_DEG = 110
      | local DISTANCE_TO_CLEARANCE = 0.300
      | local RADIUS_HELPER_POSES = 0.300
      | local RADIUS_TRANSITION_POSES = 0.400
      | local workareas = [WORKAREA_1, WORKAREA_2, WORKAREA_3, WORKAREA_4, WORKAREA_5, WORKAREA_6, WORKAREA_7, WORKAREA_8, WORKAREA_9, WORKAREA_10]
      | local poses = [PSE_WA_1, PSE_WA_2, PSE_WA_3, PSE_WA_4, PSE_WA_5, PSE_WA_6, PSE_WA_7, PSE_WA_8, PSE_WA_9, PSE_WA_10]
      | 
      | ######################### end of adjustment #########################
      | 
      | local pi = 3.14159265
      | local axis_config_current = 0
      | local axis_config_new = 0
      | local workarea_current = 0
      | local workarea_new = 0
      | global reverse_rotation = False
      | 
      | def create_translation_vector(x = 0.0, y = 0.0, z = 0.0):
      |     return struct(x = x, y = y, z = z)
      | end
      | 
      | def create_orientation_vector(rx = 0.0, ry = 0.0, rz = 0.0):
      |     return struct(rx = rx, ry = ry, rz = rz)
      | end
      | 
      | def create_transition_pose():
      |     return struct(crt = p[0,0,0,0,0,0], jnt = [0,0,0,0,0,0], q = [0,0,0,0,0,0], translation = create_translation_vector(), orientation = create_orientation_vector())
      | end
      | 
      | def compose_pose(translation = create_translation_vector(), orientation = create_orientation_vector()):
      |     return p[translation.x, translation.y, translation.z, orientation.rx, orientation.ry, orientation.rz]
      | end
      | 
      | local pose_start = create_transition_pose()
      | local pose_help = create_transition_pose()
      | local pose_target = create_transition_pose()
      | local pose = create_transition_pose()
      | 
      | def init_home_by_cartesian_pose(pose):
      |     # check given pose for reachability for the corresponding axis config
      |     local pose_home = pose_trans(pose, pose_inv(get_tcp_offset()))
      | 
      |     if check_current_axis_config() == 1:
      |         if get_inverse_kin_has_solution(pose_home, qnear=JNT_STANDARD_C1, tcp=p[0,0,0,0,0,0]):
      |             JNT_HOME = get_inverse_kin(pose_home, qnear=JNT_STANDARD_C1, tcp=p[0,0,0,0,0,0])
      |         end
      |     elif check_current_axis_config() == 2:
      |         if get_inverse_kin_has_solution(pose_home, qnear=JNT_STANDARD_C2, tcp=p[0,0,0,0,0,0]):
      |             JNT_HOME = get_inverse_kin(pose_home, qnear=JNT_STANDARD_C2, tcp=p[0,0,0,0,0,0])
      |         end
      |     end
      | end
      | 
      | def get_tool_free_pose(pose_ref=p[0,0,0,0,0,0], dir=[0,0,0], move_in_base_frame=False):
      |     # get a recovery pose
      |     # dir is providing the direction and distance in X, Y and Z
      |     # if 'move_in_base_frame' is set, dir will be interpreted as absolute values for a movement in base frame
      | 
      |     local pose_target = pose_ref
      |     local i = 0
      | 
      |     if pose_ref == p[0,0,0,0,0,0]:
      |         pose_target = get_actual_tcp_pose()
      |     end
      | 
      |     if (move_in_base_frame):
      |         while (i<3):
      |             # move only,
      |             # if the demanded position is bigger than zero and the current position is below the demanded one or
      |             # if the demanded position is smaller than zero and the current position is above the demanded one
      |             if ((dir[i]>0 and pose_target[i]<dir[i]) or (dir[i]<0 and pose_target[i]>dir[i])):
      |                 pose_target[i] = dir[i]
      |             end
      |             i = i + 1
      |         end
      |     else:
      |         pose_target = pose_trans(pose_ref, p[dir[0], dir[1], dir[2], 0, 0, 0])
      |     end
      | 
      |     return pose_target
      | end
      | 
      | def check_workarea(reference_pose):
      |     # the actual TCP position is compared to predefined areas (cubic) to determine in which area the robot arm is
      |     # a workarea is defined as a list of coordinates, where the first 3 values are X, Y, and Z with the smallest values and
      |     # the next 3 values specify X, Y and Z for the biggest values
      |     local data_size = size(workareas)
      |     local i = 0
      |     local size_workarea = p[0,0,0,0,0,0]
      |     local pose_workarea = p[0,0,0,0,0,0]
      | 
      |     while (i < data_size[0]):
      |         pose_workarea = pose_trans(inv(p[workareas[i, 0], workareas[i, 1], workareas[i, 2], 0, 0, 0]), reference_pose)
      |         size_workarea = pose_sub(p[workareas[i, 3], workareas[i, 4], workareas[i, 5], 0, 0, 0], p[workareas[i, 0], workareas[i, 1], workareas[i, 2], 0, 0, 0])
      |         if  ((pose_workarea[0]>0 and pose_workarea[0]<size_workarea[0]) and
      |             (pose_workarea[1]>0 and pose_workarea[1]<size_workarea[1]) and
      |             (pose_workarea[2]>0 and pose_workarea[2]<size_workarea[2])):
      |             return i + 1
      |         end
      |         i = i + 1
      |     end
      | 
      |     return 0
      | end
      | 
      | def check_current_axis_config():
      |     # function determnines, if the arm is oriented in one or the other configuration.
      |     # it means, that the ellbow joint is flipped and so are the wrist joints.
      | 
      |     local jnt_current = get_actual_joint_positions()
      | 
      |     # ellbow has positiv angle
      |     if (jnt_current[2]> 0):
      |         return 1
      |     # ellbow has negativ angle
      |     elif (jnt_current[2]< 0):
      |         return 2
      |     # angle is 0
      |     else:
      |         return 0
      |     end
      | end
      | 
      | def switch_axis_config(axis_config):
      |     # function to switch betwwen the axis configuration 1 and 2.
      | 
      |     if (axis_config == 1):
      |         return 2
      |     elif (axis_config ==2):
      |         return 1
      |     end
      | end
      | 
      | def get_joint_pose(pose, qnear):
      |     if get_inverse_kin_has_solution(pose, qnear=qnear):
      |         return get_inverse_kin(pose, qnear=qnear)
      |     else:
      |         popup("no solution found for the transition pose", blocking= True)
      |         return [0,0,0,0,0,0]
      |     end
      | end
      | 
      | def get_transition_pose_by_workarea(workarea):
      |     # get the correspondig pose from the list of poses
      | 
      |     pose.crt = poses[workarea-1]
      |     pose.q = set_q_near()
      |     pose.jnt = get_joint_pose(pose.crt, pose.q)
      | 
      |     return pose
      | end
      | 
      | def get_transition_pose_by_reference_pose(reference_pose, radius, keep_rxry=False):
      | 
      |     if reference_pose == p[0,0,0,0,0,0]:
      |         pose.jnt = JNT_HOME
      |         pose.q = JNT_HOME
      |         pose.crt = get_forward_kin(pose.jnt)
      |         if keep_rxry:
      |             pose.orientation = get_transition_orientation(pose.crt, keep_rxry)
      |             pose.crt = compose_pose(struct(x=pose.crt[0], y=pose.crt[1], z=pose.crt[2]), pose.orientation)
      |             pose.q = set_q_near(joints=[1,1,1,0,0,0])
      |             pose.jnt = get_joint_pose(pose.crt, pose.q)
      |         end
      |     else:
      |         pose.translation = get_transition_translation_by_radius(get_angle_to_base(reference_pose), radius)
      |         pose.orientation = get_transition_orientation(reference_pose, keep_rxry)
      |         pose.crt = compose_pose(pose.translation, pose.orientation)
      |         if keep_rxry:
      |             pose.q = set_q_near(joints=[1,1,1,0,0,0])
      |         else:
      |             pose.q = set_q_near(joints=[0,0,0,1,1,1])
      |         end
      |         pose.q[0] = adjust_axis_rotation(pose)
      |         pose.jnt = get_joint_pose(pose.crt, pose.q)
      |     end
      | 
      |     return pose
      | end
      | 
      | def get_rounded_mm(value):
      |     if (value < 0):
      |         return ceil(value*1000)
      |     elif (value >= 0):
      |         return floor(value*1000)
      |     end
      | end
      | 
      | def get_angle_to_base(pose):
      |     # get the angle relative to the base frame
      |     local pose_x_mm = 0
      |     local pose_y_mm = 0
      |     local angle = 0
      | 
      |     pose_x_mm = get_rounded_mm(pose[0])
      |     pose_y_mm = get_rounded_mm(pose[1])
      | 
      |     if (pose_x_mm == 0 and pose_y_mm < 0):
      |         angle = 0
      |     elif (pose_x_mm == 0 and pose_y_mm > 0):
      |         angle = pi
      |     elif (pose_x_mm < 0 and pose_y_mm == 0):
      |         angle = -pi/2
      |     elif (pose_x_mm > 0 and pose_y_mm == 0):
      |         angle = pi/2
      |     else:
      |         angle = atan2(pose[0], pose[1])
      |         if (-pi < angle) and (angle < 0):
      |             angle = - angle - pi
      |         elif (0 < angle) and (angle < pi):
      |             angle = - angle + pi
      |         end
      |     end
      |     return angle
      | end
      | 
      | def set_q_near(joints=[0,0,0,1,1,1], axis_config=check_current_axis_config()):
      |     local i = 0
      |     local jnt_current = get_actual_joint_positions()
      | 
      |     while i < 6:
      |         if joints[i] != 0:
      |             if axis_config == 1:
      |                 pose.q[i] = JNT_STANDARD_C1[i]
      |             elif axis_config == 2:
      |                 pose.q[i] = JNT_STANDARD_C2[i]
      |             else:
      |                 pose.q[i] = jnt_current[i]
      |             end
      |         else:
      |             pose.q[i] = jnt_current[i]
      |         end
      |         i = i + 1
      |     end
      |     return pose.q
      | end
      | 
      | def adjust_axis_rotation(pose):
      |     local angle = get_angle_to_base(pose.crt)
      | 
      |     if (0 > angle) and (angle > d2r(ANGLE_MIN_DEG)):
      |         if (pose.jnt[0] > JNT_HOME[0]):
      |             # calculated axis angle is in the wrong value range
      |             pose.q = set_q_near(joints=[1,0,0,0,0,0])
      |             reverse_rotation = True
      |         end
      |     elif (0 < angle) and (angle < d2r(ANGLE_MAX_DEG)):
      |         if (pose.jnt[0] < JNT_HOME[0]):
      |             pose.q = set_q_near(joints=[1,0,0,0,0,0])
      |             reverse_rotation = True
      |         end
      |     elif (pose.jnt[0] < -2 * pi):
      |         pose.q = set_q_near(joints=[1,0,0,0,0,0])
      |         reverse_rotation = True
      |     elif (pose.jnt[0] > 2 * pi):
      |         pose.q = set_q_near(joints=[1,0,0,0,0,0])
      |         reverse_rotation = True
      |     end
      |     return pose.q[0]
      | end
      | 
      | def get_transition_orientation(pose_ref, keep_rxry=False):
      |     # define the orientation of the transition poses
      |     local pose_current = get_actual_tcp_pose()
      |     local rpy_current = [0,0,0]
      |     local rotvec_new = [0,0,0]
      | 
      |     if keep_rxry:
      |         # use orientation of the given pose
      |         rpy_current = rotvec2rpy([pose_current[3], pose_current[4], pose_current[5]])
      |         rotvec_new = rpy2rotvec([rpy_current[0], rpy_current[1], get_angle_to_base(pose_ref) + get_locked_yaw()])
      |     else:
      |         # use orientation of defined workarea poses
      |         rpy_current = rotvec2rpy([pose_ref[3], pose_ref[4], pose_ref[5]])
      |         rotvec_new = rpy2rotvec([0, 0, rpy_current[2]])
      |     end
      |     return create_orientation_vector(rx = rotvec_new[0], ry = rotvec_new[1], rz = rotvec_new[2])
      | end
      | 
      | def get_transition_translation_by_radius(angle, radius):
      |     # calculate x,y by a radius and z by defined clearance
      |     return create_translation_vector(x = radius * cos(angle-pi/2), y = radius * sin(angle-pi/2), z = DISTANCE_TO_CLEARANCE)
      | end
      | 
      | def adjust_transition_poses(pose_identifier, keep_rxry=False):
      |     # adjust the orientation of the transition poses by determining the the current orientation
      | 
      |     local pose_current = get_actual_tcp_pose()
      |     local jnt_current = get_actual_joint_positions()
      |     local rpy_current = rotvec2rpy([pose_current[3],pose_current[4],pose_current[5]])
      |     local rotvec_new = [0,0,0]
      | 
      |     if (pose_identifier == "start"):
      |         pose = pose_start
      |     elif (pose_identifier == "target"):
      |         pose = pose_target
      |         pose.q[0] = adjust_axis_rotation(pose)
      |     elif (pose_identifier == "helper"):
      |         pose = pose_help
      |     end
      | 
      |     if keep_rxry:
      |         rotvec_new = rpy2rotvec([rpy_current[0], rpy_current[1], pose.angle_to_base + get_locked_yaw()])
      |         pose.crt = p[pose.crt[0], pose.crt[1], pose.crt[2], rotvec_new[0], rotvec_new[1], rotvec_new[2]]
      |         # adjust preferred joint angles ot the current ones
      |         pose.q[3] = jnt_current[3]
      |         pose.q[4] = jnt_current[4]
      |         pose.q[5] = jnt_current[5]
      |     end
      | 
      |     if get_inverse_kin_has_solution(pose.crt, qnear=pose.q) and is_within_safety_limits(pose.crt):
      |         pose.jnt = get_inverse_kin(pose.crt, qnear=pose.q)
      |     else:
      |         popup(str_cat("no solution for ", pose_identifier), error=True, blocking=False)
      |         pose.jnt = [0,0,0,0,0,0]
      |     end
      |     return pose.jnt
      | end
      | 
      | def get_locked_yaw():
      |     local pose_current = get_actual_tcp_pose()
      |     local rpy_current = rotvec2rpy([pose_current[3],pose_current[4],pose_current[5]])
      |     # local rotvec_new = rpy2rotvec([rpy_current[0], rpy_current[1], get_angle_to_base(pose_current)])
      |     local rotvec_new = rpy2rotvec([0, 0, get_angle_to_base(pose_current)])
      |     local pose_reference = p[pose_current[0], pose_current[1], pose_current[2], rotvec_new[0], rotvec_new[1], rotvec_new[2]]
      |     local pose_to_reference = pose_trans(pose_inv(pose_reference), pose_current)
      | 
      |     return pose_to_reference[5]
      | end
      | 
      | def get_helper_angle():
      |     local angle_start = get_angle_to_base(pose_start.crt)
      |     local angle_target = get_angle_to_base(pose_target.crt)
      |     local angle_help = (angle_start + angle_target) / 2
      | 
      |     if reverse_rotation and
      |         ((angle_start < 0 and
      |         angle_target < 0) or
      |         (angle_start > 0 and
      |         angle_target > 0)):
      |             angle_help = flip_angle(angle_help)
      |     elif (angle_start < 0 and
      |         angle_start < d2r(ANGLE_MIN_DEG)) and
      |         (angle_target > 0 and
      |         angle_target > d2r(ANGLE_MAX_DEG)):
      |             angle_help = flip_angle(angle_help)
      |     elif (angle_start > 0 and
      |         angle_start > d2r(ANGLE_MAX_DEG)) and
      |         (angle_target < 0 and
      |         angle_target < d2r(ANGLE_MIN_DEG)):
      |             angle_help = flip_angle(angle_help)
      |     end
      |     return angle_help
      | end
      | 
      | def flip_angle(angle):
      |     # flips the given angle 180 degree around
      |     if (angle < 0):
      |         return angle + pi
      |     elif (angle > 0):
      |         return angle - pi
      |     end
      | end
      | 
      | def clear_poses():
      |     pose = create_transition_pose()
      |     pose_start = create_transition_pose()
      |     pose_help = create_transition_pose()
      |     pose_target = create_transition_pose()
      | end
      | 
      | def do_transition(reference_pose=p[0,0,0,0,0,0], mode=2, keep_rxry=False, a=1.4, v=1.05, r=0.100):
      |     # the robot will evaluate the current and target workarea
      |     # after that, the robot will move between the workareas automatically.
      |     # parameters:
      |     # reference_pose:   a pose/frame were the robot should work next. If nothing is given, base frame will be used as target
      |     # keep_rxry:        if true, the robot will keep the orientation of the tool during the movement
      | 
      |     ################# checking #################
      |     clear_poses()
      |     workarea_current = check_workarea(get_actual_tcp_pose())    # between 0 and the amount of defined workareas
      |     workarea_new = check_workarea(reference_pose)               # between 0 and the amount of defined workareas
      |     reverse_rotation = False
      | 
      |     if (workarea_current != 0 and workarea_new != 0 and workarea_current != workarea_new) or (reference_pose == p[0,0,0,0,0,0]):
      |         ################# get axisvalues #################
      |         if (mode == 1):
      |             pose_start = get_transition_pose_by_workarea(workarea_current)
      |             pose_target = get_transition_pose_by_workarea(workarea_new)
      |         elif (mode == 2):
      |             pose_start = get_transition_pose_by_reference_pose(get_actual_tcp_pose(), RADIUS_TRANSITION_POSES, keep_rxry)
      |             pose_target = get_transition_pose_by_reference_pose(reference_pose, RADIUS_TRANSITION_POSES, keep_rxry)
      | 
      |         end
      |         # if (pose_start.crt[1] < 0 and pose_target.crt[1] > 0) or (pose_start.crt[1] > 0 and pose_target.crt[1] < 0):
      |         #     pose_help = get_transition_pose_by_reference_pose(pose_start.crt, RADIUS_HELPER_POSES)
      |         # end
      |         textmsg("Cartesian pose start: ", to_str(pose_start.crt))
      |         textmsg("Joints pose start: ", to_str(pose_start.jnt))
      |         textmsg("Qnear pose start: ", to_str(pose_start.q))
      |         textmsg("Cartesian pose target: ", to_str(pose_target.crt))
      |         textmsg("Joints pose target: ", to_str(pose_target.jnt))
      |         textmsg("Qnear pose target: ", to_str(pose_target.q))
      | 
      |         ################# movements #################
      |         if (pose_help.jnt != [0,0,0,0,0,0]):
      |             if point_dist(get_actual_tcp_pose(), pose_start.crt) > r and point_dist(pose_start.crt, pose_help.crt) > r:
      |                 movej(pose_start.jnt, a=a, v=v, r=r)
      |                 if (point_dist(pose_start.crt, pose_help.crt) > r) and (point_dist(pose_target.crt, pose_help.crt) > r):
      |                     movej(pose_help.jnt, a=a, v=v, r=r)
      |                 end
      |             end
      |         else:
      |             if point_dist(get_actual_tcp_pose(), pose_start.crt) > r and point_dist(pose_start.crt, pose_target.crt) > r:
      |                 movej(pose_start.jnt, a=a, v=v, r=r)
      |             end
      |         end
      |         movej(pose_target.jnt, a=a, v=v)
      | 
      |         ################# checking #################
      |         workarea_current = check_workarea(get_actual_tcp_pose())    # between 0 and the amount of defined workareas
      |     else:
      |         # define error or warning
      |     end
      | end
      | 
      | 
      | # Erläuterung
      | # für start wird die aktuelle Position übergeben
      | # davon wird die Position für start berechnet. Bei der Orientierung wird entweder nur Rz genommen oder alles bei keep_rxry
    Script file /programs/04 Scripts/SCRIPT Logs V1.2.script
      | current_state_log = ""
      | current_process_log = ""
      | current_step_log = ""
      | current_warning_log = ""
      | current_error_log = ""
      | current_hatch_log = ""
      | current_centrifuge_log = ""
      | current_message_log = "placeholderstring"
      | LogLevel=struct(NONE=0, INFO=1, PROCESS=2, WARNING=3, ERROR=4)
      | LOGLEVEL=LogLevel.INFO
      | 
      | def log_message(prefix="", newlog=current_message_log):
      |     # generates a log message every time its useful
      |     if (current_message_log != newlog and newlog != ""):
      |         textmsg(str_cat(prefix, to_str(newlog)))
      |         current_message_log = to_str(newlog)
      |     end
      | end
      | 
      | def log_state(newlog):
      |     # generates a log message every time its useful
      |     if (current_state_log != newlog and newlog != ""):
      |         textmsg(str_cat("Machine: ", to_str(newlog)))
      |         current_state_log = to_str(newlog)
      |     end
      | end
      | 
      | def log_process(newlog):
      |     # generates a log message every time its useful
      |     if (current_process_log != newlog and newlog != ""):
      |         textmsg(str_cat("Process: ", to_str(newlog)))
      |         current_process_log = to_str(newlog)
      |     end
      | end
      | 
      | def log_step(newlog):
      |     # generates a log message every time its useful
      |     if (current_step_log != newlog and newlog != ""):
      |         textmsg(str_cat("Step: ", to_str(newlog)))
      |         current_step_log = to_str(newlog)
      |     end
      | end
      | 
      | def log_info(newlog):
      |     # generates a log message if log level is Info or lower
      |     if (newlog != "" and LOGLEVEL <= LogLevel.INFO):
      |         textmsg(str_cat("INFO: ", newlog))
      |     end
      | end
      | 
      | def log_warning(newlog):
      |     # generates a log message every time its useful
      |     if (current_warning_log != newlog and newlog != ""):
      |         textmsg(str_cat("WARNING: ", to_str(newlog)))
      |         current_warning_log = to_str(newlog)
      |     end
      | end
      | 
      | def log_error(newlog):
      |     # generates a log message every time its useful
      |     if (current_error_log != newlog and newlog != ""):
      |         textmsg(str_cat("ERROR: ", to_str(newlog)))
      |         current_error_log = to_str(newlog)
      |     end
      | end
      | 
      | def log_hatch_state(newlog):
      |     # generates a log message every time its useful
      |     if (current_hatch_log != to_str(newlog) and to_str(newlog) != ""):
      |         textmsg(str_cat("Hatch_state: ", to_str(newlog)))
      |         current_hatch_log = to_str(newlog)
      |     end
      | end
      | 
      | def log_centrifuge_state(newlog):
      |     # generates a log message every time its useful
      |     if (current_centrifuge_log != to_str(newlog) and to_str(newlog) != ""):
      |         textmsg(str_cat("Centrifuge_state: ", to_str(newlog)))
      |         current_centrifuge_log = to_str(newlog)
      |     end
      | end
    Script file /programs/04 Scripts/SCRIPT Statistics V1.1.script
      | #*****************************************************
      | # customer          :   tbd
      | # project name      :   tbd
      | #****************************************************
      | # controller        :
      | # software          :
      | #****************************************************
      | # author            :   P. Koehnke (+49 1628859904; p.koehnke@unitedrobotics.group)
      | # Copyright (c)     :   United Robotics Group Health and Food GmbH
      | #                       An der Riede 2
      | #                       28816 Stuhr
      | #                       Germany
      | #****************************************************
      | # description       :   statistics script, which tracks the times in different PackML states and let you count objects
      | # version:      	:   1.0
      | # created           :   20.11.2023
      | # updated           :
      | #****************************************************
      | # modifications     :
      | #
      | # date              :
      | # name              :
      | # reason            :
      | #****************************************************
      | 
      | # to save the times persistently, these variables must be defined in the installation file of the robot
      | 
      | # ===== object counters =====
      | def count_up(counters, idx, by):
      |     counters[idx] = counters[idx] + by
      |     return counters
      | end
      | 
      | def count_total(counters):
      |     local i = 0
      |     local total = 0
      |     while (i<length(counters)):
      |         total = total + counters[i]
      |         i = i + 1
      |     end
      |     return total
      | end
      | # ==========
      | 
      | # ===== Times =====
      | thread Pml_Timer_Thread():
      |     # STATE_Times is a list of all time values in seconds
      |     while (True):
      |         STATE_Times[STATE-1] = STATE_Times[STATE-1] + get_steptime()
      |         sync()
      |     end
      | end
      | 
      | thread_timer_handler = run Pml_Timer_Thread()
      | 
      | def get_time(timer, format="dd/hh/mm/ss"):
      |     # give the time in seconds
      |     # the function will return the given time as string in the predefined format
      |     local days = floor(timer/86400)
      |     local hours = floor((timer%86400)/3600)
      |     local minutes = floor((timer%3600)/60)
      |     local seconds = floor(timer%60)
      |     return str_cat(str_cat(str_cat(str_cat(str_cat(str_cat(to_str(days), "/"), to_str(hours)), "/"), to_str(minutes)), "/"), to_str(seconds))
      | end
      | 
      | def set_timer(time, format="dd/hh/mm/ss"):
      |     # give the time as string
      |     # the function will return the corresponding seconds summed up
      |     local days_idx = str_find(time, "/", 0)
      |     local hours_idx = str_find(time, "/", days_idx+1)
      |     local minutes_idx = str_find(time, "/", hours_idx+1)
      |     local days = to_num(str_sub(time, 0, days_idx))
      |     local hours = to_num(str_sub(time, days_idx+1, hours_idx-days_idx-1))
      |     local minutes = to_num(str_sub(time, hours_idx+1, minutes_idx-hours_idx-1))
      |     local seconds = to_num(str_sub(time, minutes_idx+1, length(time)-minutes_idx))
      |     return (days*86400 + hours*3600 + minutes*60 + seconds)
      | end
    Script file /programs/04 Scripts/SCRIPT Vision Config V0.2.script
      | CAM_LM = struct(id=0, type="", size=0, related_itm=0, capture_relation="")
      | global CAM_Result = make_list(0, 0, 50)
      | 
      | def create_landmark(id=0, type="", size=0, related_itm=0, capture_relation=""):
      |     return struct(id=id, type=type, size=size, related_itm=related_itm, capture_relation=capture_relation)
      | end
      | 
      | 
      | CAM_LMs = [
      |   create_landmark(id=1, type="aruco_7x7", size=0.1, related_itm=1, capture_relation="front_right"),
      |   create_landmark(id=4, type="aruco_7x7", size=0.1, related_itm=2, capture_relation="straight_left"),
      |   create_landmark(id=3, type="aruco_7x7", size=0.1, related_itm=2, capture_relation="straight_left"),
      |   create_landmark(id=8, type="aruco_7x7", size=0.1, related_itm=2, capture_relation="right"),
      |   create_landmark(id=5, type="aruco_7x7", size=0.1, related_itm=5, capture_relation="left"),
      |   create_landmark(id=6, type="aruco_7x7", size=0.1, related_itm=2, capture_relation="straight_left")
      | ]
      | 
      | CAM_Capture_Poses = struct(
      |   front_left = p[0.350,-0.330,0.500,0.353,-0.323,-1.458],
      |   left = p[0.350,0.000,0.500,0.353,-0.323,-1.458],
      |   back_left = p[0.350,0.220,0.500,0.353,-0.323,-1.458],
      |   back_right = p[-0.350,0.000,0.500,0.579,0.240,0.760],
      |   right = p[-0.350,-0.300,0.500,0.206,0.206,1.561],
      |   front_right = p[-0.350,-0.400,0.500,0.242,0.903,2.480],
      |   straight_left = p[0.375,-0.000,0.500,0.815,-0.815,-1.412],
      |   front = p[0,0,0,0,0,0]
      | )
      | 
      | def get_capture_pose(lm):
      |     if (lm.capture_relation == "front_left"):
      |         return CAM_Capture_Poses.front_left
      |     elif (lm.capture_relation == "left"):
      |         return CAM_Capture_Poses.left
      |     elif (lm.capture_relation == "back_left"):
      |         return CAM_Capture_Poses.back_left
      |     elif (lm.capture_relation == "back_right"):
      |         return CAM_Capture_Poses.back_right
      |     elif (lm.capture_relation == "right"):
      |         return CAM_Capture_Poses.right
      |     elif (lm.capture_relation == "straight_left"):
      |        return CAM_Capture_Poses.straight_left
      |     else:
      |         # error
      |         return get_actual_tcp_pose()
      |     end
      | end
    Script file /programs/04 Scripts/SCRIPT uLM Factory.script
      | # ############### SCRIPT uLM Factory ##################
      | # *****************************************************
      | # Customer          :   URG
      | # Product Name      :   uLabMobile
      | # ****************************************************
      | # Controller/Robot  :   UR5e
      | # Software          :   URSCRIPT
      | # Dependencies      :   Defines Script but mainly independend
      | # How To            :   is used by projectconfig to create list of structs full of projectrelated information which are used across the scripts
      | # ****************************************************
      | # Author            :   D.Kreugel
      | # Copyright (c)     :   United Robotics Group Health and Food GmbH
      | #                       An der Riede 2
      | #                       28816 Stuhr
      | #                       Germany
      | # ****************************************************
      | # Description       :   definition of the datastructures used by the uLM, gives functionality to create a predefined datastructure, is assigned to a global list in projectconfig
      | # Version           :   0.2
      | # Created           :   18.07.2024
      | # Updated           :
      | # ****************************************************
      | # Modifications     :
      | #
      | # Date              :
      | # Name              :
      | # Reason            :
      | # ****************************************************
      | # TODO              : cleanup useless info and add all other factorys from the other scripts here to have one place to search for such things, documentation
      | 
      | # DO NOT TOUCH THE DATASTRUCTURES IF YOU DON'T KNOW WHAT YOU DO!
      | MAX_ACTIONS=6
      | POS_Z=p[0,0,0,0,0,0]
      | def create_pattern(id=0, name="", pattern_width=[0, 0], pattern_size=[0, 0], blocked=[-1, -1, -1], direction="X", transpose=False, invert=False, description="default"):
      |     return struct(
      |         id = id,
      |         name = name,
      |         pattern_width = pattern_width,
      |         pattern_size = pattern_size,
      |         blocked = blocked,
      |         direction = direction,
      |         transpose = transpose,
      |         invert = invert,
      |         description = description
      |     )
      | end
      | 
      | # item model stores frame related inner and outer patterns
      | def create_item_model(inner="", outer="", description="default"):
      |     return struct(
      |         inner = inner,
      |         outer = outer,
      |         description = description
      |         )
      | end
      | 
      | # creates a fixed length list cause structs cannot deal with dynamic lists at the moment and an item can have different amount of actions assigned to it
      | def create_action_list(values):
      |     local list = make_list(MAX_ACTIONS, 0, MAX_ACTIONS+1)
      |     local i = 0
      |     while (i < values.length()):
      |         list[i] = values[i]
      |         i = i + 1
      |     end
      |     return list
      | end
      | 
      | def create_item(id=0, ls_item="default", frame=p[0,0,0,0,0,0], actionlist=create_action_list([]), item_model=create_item_model(), lm_id=0, description="default"):
      |     return struct(
      |         id = id,
      |         ls_item = ls_item,
      |         frame = frame,
      |         actionlist = create_action_list(actionlist),
      |         item_model = item_model,
      |         lm_id = lm_id,
      |         description = description
      |     )
      | end
      | 
      | def create_object(id=0, obj_name=0, height=0, width=0, obj_type = 0, description="default"):
      |     return struct(
      |         id = id,
      |         obj_name = obj_name,
      |         obj_type = obj_type,
      |         height = height,
      |         width = width,
      |         description = description
      |     )
      | end
      | # extends object type by sample related information
      | def create_sample(obj_id=0, cap_diameter=0, raw_diameter=0, color="", material="", description=""):
      |     return struct(
      |     obj_id = obj_id,
      |     cap_diameter = cap_diameter,
      |     raw_diameter = raw_diameter,
      |     color = color,
      |     material = material,
      |     description = description)
      | end
      | 
      | # create gripper configs
      | def create_gripper_config(gripper_offset=struct(prepick=2, pick=0, place=2), force=0, speed=0, validation=0, object=create_object()):
      |     gripper_offset.prepick = object.width+gripper_offset.prepick
      |     gripper_offset.place = object.width+gripper_offset.place
      |     return struct(
      |         object = object.obj_name,
      |         force = force,
      |         speed = speed,
      |         validation = validation,
      |         width = gripper_offset
      |     )
      | end
      | 
      | def create_manipulator_command(id="", item="", action=0, jig_nbr=-1, obj_nbr=-1, object_type=-1, error_id=0, data=""):
      |     return struct(
      |         id = id,
      |         device = Device.MANIPULATOR,
      |         item = item,
      |         action = action,
      |         jig_nbr = jig_nbr,
      |         obj_nbr = obj_nbr,
      |         object_type = object_type,
      |         error_id = error_id,
      |         data = data
      |     )
      | end
      | 
      | def create_amr_command(id="", item="", action=0, target=0, error_id=0, data=""):
      |     return struct(
      |         id = id,
      |         device = Device.AMR,
      |         item = item,
      |         action = action,
      |         target = target,
      |         error_id = error_id,
      |         data = data
      |     )
      | end
      | 
      | def create_camera_command(id="", item="", action=0, attempt=0, error_id=0, data=""):
      |     return struct(
      |         id = id,
      |         device = Device.CAMERA,
      |         item = item,
      |         action = action,
      |         attempt = attempt,
      |         error_id = error_id,
      |         data = data
      |     )
      | end
      | 
      | # Function to create a new  vision struct to assign workspace and skill to an item or a selection
      | def create_vision_config(workspace_id="", skill_id="", item_id=-1, target_origin=p[0,0,0,0,0,0], description="default"):
      |     return struct(
      |         workspace_id = workspace_id,
      |         skill_id = skill_id,
      |         item_id = item_id,
      |         target_origin = target_origin,
      |         description = description)
      | end
      | 
      | # extents the vision config by the inspect configuration, this info will be called in the action inspect only
      | # item_id is the reference to the item
      | # dx is the distance in x direction for one position to the next in the inspection rack
      | # dy is the distance in y direction for one position to the next in the inspection rack
      | # target origin is the origin coordinate of the first position in the inspectionrack from where the calculation starts
      | def create_inspect_config(item_id=0, dx=0, dy=0, target_origin=p[0,0,0,0,0,0], rack_size=[0,0], description="default"):
      |     return struct(
      |     item_id = item_id,
      |     dx = dx,
      |     dy = dy,
      |     target_origin = target_origin,
      |     rack_size = rack_size,
      |     description = description
      |     )
      | end
      |  # Function to create a new landmark struct that contains all lm related configurationparameters and will be assigned via item_id
      | #def create_landmark(lm_id=0, marker_id=-1, marker_size=0.1, marker_type="aruco_7x7", capture_pos=p[0,0,0,0,0,0], init_frame=p[0,0,0,0,0,0], search_offset=[0,0,0], actual_frame=p[0,0,0,0,0,0], description=""):
      |   ##  return struct(
      |    #     lm_id = lm_id,
      |    #     marker_id = marker_id,
      |      #   marker_size = marker_size,
      |   ##      marker_type = marker_type,
      |   #      capture_pos = capture_pos,
      |   #      init_frame = init_frame,
      |   #      search_offset = search_offset,
      |   #      actual_frame = actual_frame,
      | #        description = description)
      | #end
      | 
      | def create_movement(id=0, actionlist=create_action_list([]), hh_approach=POS_Z, h_approach=POS_Z, approach=POS_Z, h_target=POS_Z, target=POS_Z, retract=POS_Z, h_retract=POS_Z, hh_retract=POS_Z, h_frame=POS_Z, frame=POS_Z, speed=1, acceleration=1, description="default"):
      | return struct(
      |     id = id,
      |     actionlist = actionlist,
      |     hh_approach = hh_approach,
      |     h_approach = h_approach,
      |     approach = approach,
      |     h_target = h_target,
      |     target = target,
      |     retract = retract,
      |     h_retract = h_retract,
      |     hh_retract = hh_retract,
      |     h_frame = h_frame,
      |     frame = frame,
      |     speed = speed,
      |     acceleration = acceleration,
      |     description = description
      | )
      | end
    Script file /programs/04 Scripts/SCRIPT uLM Defines v0.2.script
      | ############# SCRIPT uLM Defines ###############
      | #*****************************************************
      | # Customer          :   URG
      | # Product Name      :   uLabMobile
      | #****************************************************
      | # Controller/Robot  :   UR5e
      | # Software          :   5.17
      | # Dependencies      :   Factory Script, Logs Script
      | # How To            :   Define Constants depending on the Project, don't go to big in Listsize as it will exceed the URScript limits
      | #****************************************************
      | # Author            :   D.Kreugel
      | # Copyright (c)     :   United Robotics Group Health and Food GmbH
      | #                       An der Riede 2
      | #                       28816 Stuhr
      | #                       Germany
      | #****************************************************
      | # Description       :   Defines all Enums and Global reachable Varibles/Datastructures
      | # Version           :   0.2
      | # Created           :   18.07.2024
      | # Updated           :
      | #****************************************************
      | # Modifications     :
      | #
      | # Date              :
      | # Name              :
      | # Reason            :
      | #****************************************************
      | # TODO find better place for the Search Funktions for the Object Lists, documentation
      | 
      | 
      | POS_Z = p[0,0,0,0,0,0]
      | 
      | # DEFAULTS ROBOT MOVEMENTS
      | DEFAULT = struct(SPEED=0.8, ACCELERATION=0.6)
      | 
      | # ENUMS
      | Objects = struct(NONE=0, CC_SAMPLE=1, CC_RACK=2, COAG_SAMPLE=3, COAG_RACK=4, HEMA_SAMPLE=5, HEMA_RACK=6, INPUT_RACK=7, CF_RACK=8, ANY_SAMPLE=9, ANY_RACK=10, TARA_SAMPLE=11, BUTTON=12, XN550_DRAWER=13, COBAS_RACK=14)
      | ObjectType = struct(NONE=0,SAMPLE=1,RACK=2, BUTTON=3, DRAWER=4)
      | 
      | ActionManipulator = struct(NONE=0, PICK=1, PLACE=2, DECAP=12, PUSH=3, RELEASE=21, GRASP=20, MOVE_TO=19, DRAWER_OPEN=51, DRAWER_CLOSE=52)
      | ActionAMR = struct(NONE=0, LOAD_MISSION=31, START_MISSION=32, NAVIGATE=33, ACKNOWLEDGE=34, READ=35)
      | ActionCamera = struct(NONE=0, INSPECT=16, DETECT=15, DETECT_OBJECTS=17)
      | Device = struct(MANIPULATOR=1, AMR=2, CAMERA=3)
      | Patterns = struct(NONE="NONE", TARA="TARA", CENTRIFUGE="CENTRIFUGE",CENTRIFUGE_MAGAZINE="CENTRIFUGE_MAGAZINE",SYSMEX_XN550="SYSMEX_XN550",COBAS="COBAS",COBAS_MAGAZINE="COBAS_MAGAZINE",INPUT="INPUT",NOK="NOK",DRAWER_XN550="DRAWER_XN550",ARCHIVE="ARCHIVE")
      | CommandStatus = struct(EXECUTED=0, UNFINISHED=1)
      | 
      | # Constants
      | MAX_CAPTURE_ATTEMPTS = 8
      | # Maximum Size of the Datastructures
      | MAX_ITEM_OBJ = 40
      | MAX_GRIPPER_OBJ = 10
      | MAX_LANDMARK_OBJ = 10
      | MAX_PATTERN_OBJ = 30
      | MAX_ITEM_MODEL_OBJ = 20
      | MAX_VISION_CONFIG_OBJ = 10
      | MAX_CAPTURE_RESULTS = 55
      | MAX_MOVEMENT_OBJ = 50
      | 
      | CON=False
      | 
      | # for Marburg Approach
      | LAST_CAPTURE = make_list(0, "", MAX_CAPTURE_RESULTS)
      | 
      | # Initialize the Datastructures in order to store related Data and use them in structs without length issues
      | 
      | OBJECT_MAP = make_list(0 ,create_object(), MAX_ITEM_OBJ)
      | ITEM_MAP = make_list(0, create_item(), MAX_ITEM_OBJ)
      | ITEM_MODEL_MAP = make_list(0, create_pattern(), MAX_ITEM_MODEL_OBJ)
      | GRIPPER_CONFIG_MAP = make_list(0, create_gripper_config(), MAX_PATTERN_OBJ)
      | VISION_CONFIG_MAP = make_list(0, create_vision_config(), MAX_VISION_CONFIG_OBJ)
      | INSPECT_CONFIG_MAP = make_list(0, create_inspect_config(), MAX_VISION_CONFIG_OBJ)
      | LANDMARK_MAP = make_list(0, create_landmark(), MAX_LANDMARK_OBJ)
      | MOVEMENT_MAP = make_list(0, create_movement(), MAX_MOVEMENT_OBJ)
      | 
      | OBJECT_REFERENCE_HEIGHT = 81
      | 
      | 
      | # functions to search in the datastructures which are defined in the factories
      | 
      | ################# MOVEMENT ###############
      | 
      | def find_movement_by_frame_and_action(frame,action):
      |     local i = 0
      |     local ii = 0
      |     while (i < MOVEMENT_MAP.length()):
      |         if (MOVEMENT_MAP[i].frame == frame):
      |             while(ii < MOVEMENT_MAP[i].actionlist.length()):
      |                 if (MOVEMENT_MAP[i].actionlist[ii] == action):
      |                     log_info("Movement found: [" + to_str(MOVEMENT_MAP[i].description) + "]")
      |                     return MOVEMENT_MAP[i]
      |                 end
      |                 ii = ii + 1
      |             end
      |             ii = 0
      |         end
      |         i = i + 1
      |     end
      |     log_warning("no movement found for frame: [" + to_str(frame) + "]")
      |     return create_movement(frame=frame)  # Return default pattern if not found
      | end
      | 
      | def find_item_by_lsitem_and_action(ls_item, action):
      |     local i = 0
      |     while (i < ITEM_MAP.length()):
      |         if (ITEM_MAP[i].ls_item == ls_item):
      |             local ii = 0
      |             while (ii < ITEM_MAP[i].actionlist.length()):
      |                 if (ITEM_MAP[i].actionlist[ii] == action):
      |                     log_info("Item found: [" + to_str(ITEM_MAP[i].description) + "]")
      |                     return ITEM_MAP[i]
      |                 end
      |                 ii = ii + 1
      |             end
      |         end
      |         i = i + 1
      |     end
      |     log_warning("Item not found for station[" + to_str(ls_item) + "] and action[" + to_str(action) + "]")
      |     return create_item()  # Return default item if not found
      | end
      | ################# PATTERN ###################
      | 
      | def find_pattern_by_name(name):
      |     local i = 0
      |     while (i < ITEM_MODEL_MAP.length()):
      |         if (ITEM_MODEL_MAP[i].name == name):
      |             log_info("Item Model found: [" + to_str(ITEM_MODEL_MAP[i].description) + "]")
      |             return ITEM_MODEL_MAP[i]
      |         end
      |         i = i + 1
      |     end
      |     log_warning("Item Model not found for name[" + to_str(name) + "]")
      |     return create_pattern()  # Return default pattern if not found
      | end
      | 
      | def is_in_list(list,val):
      |     local i = 0
      |     while(i<list.length()):
      |         if(list[i]==val):
      |             return True
      |         end
      |         i=i+1
      |     end
      |     return False
      | end
      | 
      | def get_next_valid_patternslot(item_model, counter):
      |     local i = 0
      |     local temp = 0
      |     local max_slots = item_model.pattern_size[0] * item_model.pattern_size[1]
      |     log_info("blocked positions:" + to_str(item_model.blocked) + "| current pos: " + to_str(counter))
      |     while (i < item_model.blocked.length()):
      |         if(item_model.blocked[i] <= counter and item_model.blocked[i] != -1):
      |             temp = temp + 1
      |         end
      |         i = i + 1
      |     end
      | 
      |     if(is_in_list(item_model.blocked,counter+temp)):
      |         while(is_in_list(item_model.blocked,counter+temp)):
      |             temp=temp+1
      |         end
      |     end
